Fanuc KAREL source: kc00033.KL

PROGRAM KC00033
%STACKSIZE=65535
%PRIORITY=65535
%NOLOCKGROUP
VAR
I : INTEGER
J : INTEGER
K : INTEGER
R : REAL
B : BOOLEAN
S : STRING[80]
T : STRING[80]
AI : ARRAY[8] OF INTEGER
AB : ARRAY[244] OF BYTE
JP : JOINTPOS9
AR : ARRAY[6] OF REAL
-- UNRESOLVED DECLARATIONS (source type spelling not recovered)
-- P : TYPE_0x001F (type_u16=0x001F)
-- Q : TYPE_0x001F (type_u16=0x001F)
BEGIN
-- UNRESOLVED_PC line 18 opcodes [27 22 1C 22 22 76] marker_code=0
END KC00033
